Fanuc KAREL source: KC00020.KL

PROGRAM KC00020
%NOLOCKGROUP
%ENVIRONMENT MOTN
VAR
  I: INTEGER
  J: INTEGER
  K: INTEGER
  R: REAL
  B: BOOLEAN
  S: STRING[80]
  T: STRING[80]
  P: PATH
  Q: PATH
  AI: ARRAY[8] OF INTEGER
  AB: ARRAY[244] OF BYTE
BEGIN
  CNCL_STP_MTN
END KC00020
